// TIA Portal V21 export
// export: Created 2026-11-22T02:34:23.1888706Z, ExportSetting WithDefaults, DisplayName Totally Integrated Automation Portal, DisplayVersion V21 Update 3, DisplayName STEP 7 Professional, DisplayVersion V21 Update 3, DisplayName STEP 7 Safety, DisplayVersion V21, DisplayName Tech WebApplication, DisplayVersion V21, DisplayName WinCC Basic/Comfort/Advanced, DisplayVersion V21 Update 3, DisplayName WinCC Unified, DisplayVersion V21 Update 3
TextList "TL_BitNo"  ListRange=Binary
  TextListEntry   EntryType=SingleValue, Text="Bit 0 set"
  TextListEntry   EntryType=SingleValue, From=1, To=1, Text="Bit 1 set"
  TextListEntry   EntryType=SingleValue, From=2, To=2, Text="Bit 2 set"
  TextListEntry   EntryType=SingleValue, From=3, To=3, Text="Bit 3 set"
